// TIA Portal project "FillingLine" (V21)

(* hardware
DEVICE "PLC_Line"  S7-1500 station
   slot 0: "Rail_0"  Rack  6ES7 590-1***0-0AA0
   slot 1: "PLC_Line"  CPU 1516-3 PN/DP  6ES7 516-3AN02-0AB0  V2.9
      slot 3: "CPU display_1"  6ES7591-1BA00-0AA0
      slot 32768: "PROFINET interface_1"  X1
         slot 32769: "Port_1"  X1 P1
         slot 32770: "Port_2"  X1 P2
      slot 33024: "PROFINET interface_2"  X2
         slot 33025: "Port_1"  X2 P1
      slot 33280: "DP interface_1"  X3
      slot 34817: "Virtual CP interface port_1"  Virtual CP interface port  Virtual CP interface port
*)

// ===== PLC "PLC_Line"  CPU 1516-3 PN/DP =====

VAR_GLOBAL   // PLC tag table "Inputs"
   "Button_Start" AT %I0.0 : Bool;   // Start the line
   "Button_Stop" AT %I0.1 : Bool;   // Stop the line, normally closed
   "Button_Reset" AT %I0.2 : Bool;   // Acknowledge faults
   "Infeed_BottleAtFiller" AT %I1.0 : Bool;   // Photo eye: a bottle stands under the filler
   "Infeed_MotorFeedback" AT %I1.1 : Bool;   // Infeed contactor is closed
   "Outfeed_BottleAtEnd" AT %I1.2 : Bool;   // Photo eye at the end of the outfeed
   "Outfeed_MotorFeedback" AT %I1.3 : Bool;   // Outfeed contactor is closed
   "Filler_ValveOpened" AT %I1.4 : Bool;   // Fill valve is open
   "Filler_ValveClosed" AT %I1.5 : Bool;   // Fill valve is closed
   "Packer_Ready" AT %I1.6 : Bool;   // The packer can take a bottle
   "Filler_Level" AT %IW64 : Int;   // Level in the bottle, raw 0 to 27648
END_VAR

VAR_GLOBAL   // PLC tag table "Operator"
   "Recipe_Selected" AT %MW10 : Int;   // Recipe chosen on the panel, 1 to 3
   "Bottles_Filled" AT %MD12 : DInt;   // Bottles filled since the last start
END_VAR

VAR_GLOBAL   // PLC tag table "Outputs"
   "Infeed_Motor" AT %Q0.0 : Bool;   // Infeed conveyor motor
   "Outfeed_Motor" AT %Q0.1 : Bool;   // Outfeed conveyor motor
   "Filler_Valve" AT %Q0.2 : Bool;   // Opens the fill valve
   "Lamp_Running" AT %Q0.3 : Bool;   // The line runs
   "Lamp_Fault" AT %Q0.4 : Bool;   // A fault waits to be acknowledged
END_VAR

// folder: Line

TYPE "typeRecipe"
   STRUCT
      label : String[20];   // Shown on the panel
      volume : Real;   // Fill volume in ml
      settleTime : Time;   // Foam settles before the bottle moves on
   END_STRUCT;
END_TYPE

// folder: Data

DATA_BLOCK "Recipes"   // DB1
{ S7_Optimized_Access := 'TRUE' }
VERSION : 0.1
   VAR
      active : "typeRecipe";   // The recipe in use
      list : Array[1..3] of "typeRecipe";   // Recipes to choose from
   END_VAR
BEGIN
   list[1].label := 'Water 0.5 l';
   list[1].volume := 500.0;
   list[1].settleTime := T#500MS;
   list[2].label := 'Water 1 l';
   list[2].volume := 1000.0;
   list[2].settleTime := T#800MS;
   list[3].label := 'Soda 0.5 l';
   list[3].volume := 480.0;
   list[3].settleTime := T#3S;
END_DATA_BLOCK

DATA_BLOCK "LineData"   // DB2
{ S7_Optimized_Access := 'TRUE' }
VERSION : 0.1
// stored: InstanceOfName FillingLine
"FillingLine"
BEGIN
END_DATA_BLOCK

// folder: (top level)

ORGANIZATION_BLOCK "Main"   // OB1, SCL, ProgramCycle
TITLE = "Main Program Sweep (Cycle)"
{ S7_Optimized_Access := 'TRUE' }
VERSION : 0.1
   VAR_INPUT
      Initial_Call : Bool;   // Initial call of this OB
      Remanence : Bool;   // =True, if remanent data are available
   END_VAR
BEGIN

    // Take the recipe the operator chose, then run the line.
    "Recipes".active := "Recipes".list[LIMIT(MN := 1, IN := "Recipe_Selected", MX := 3)];

    "LineData"(start := "Button_Start",
               stop := NOT "Button_Stop",
               reset := "Button_Reset");

    "Lamp_Running" := "LineData".running;
    "Lamp_Fault" := "LineData".fault;
END_ORGANIZATION_BLOCK

// folder: Common

FUNCTION_BLOCK "Motor"   // FB1, SCL
TITLE = Motor with feedback
{ S7_Optimized_Access := 'TRUE' }
VERSION : 0.1
// Starts and stops a motor and watches its contactor's feedback.
   VAR_INPUT
      start : Bool;   // Start command
      stop : Bool;   // Stop command, wins over start
      feedback : Bool;   // Contactor is closed
      reset : Bool;   // Acknowledge a fault
   END_VAR
   VAR_OUTPUT
      run : Bool;   // Drives the contactor
      fault : Bool;   // The feedback did not come in time
   END_VAR
   VAR
      feedbackTimer : TON_TIME;
      enabled : Bool;   // Started and not stopped since
   END_VAR
   VAR CONSTANT
      FEEDBACK_TIME : Time := T#2S;   // How long the contactor may take
   END_VAR
BEGIN

    // Stop wins over start, and a fault keeps the motor off until it is reset.
    IF #stop OR #fault THEN
        #enabled := FALSE;
    ELSIF #start THEN
        #enabled := TRUE;
    END_IF;

    #feedbackTimer(IN := #enabled AND NOT #feedback,
                   PT := #FEEDBACK_TIME);
    IF #feedbackTimer.Q THEN
        #fault := TRUE;
    ELSIF #reset THEN
        #fault := FALSE;
    END_IF;

    #run := #enabled AND NOT #fault;
END_FUNCTION_BLOCK

FUNCTION_BLOCK "Valve"   // FB2, SCL
TITLE = Valve with end switches
{ S7_Optimized_Access := 'TRUE' }
VERSION : 0.1
// Opens and closes a valve and checks that it reaches its end position in time.
   VAR_INPUT
      open : Bool;   // Open the valve
      opened : Bool;   // End switch: open
      closed : Bool;   // End switch: closed
      reset : Bool;   // Acknowledge a fault
   END_VAR
   VAR_OUTPUT
      output : Bool;   // Drives the valve
      fault : Bool;   // An end position was not reached in time
   END_VAR
   VAR
      moveTimer : TON_TIME;
   END_VAR
   VAR CONSTANT
      MOVE_TIME : Time := T#1S;   // How long the valve may take to move
   END_VAR
BEGIN

    #output := #open AND NOT #fault;

    // The valve is moving while it is not where it was told to go.
    #moveTimer(IN := (#output AND NOT #opened) OR (NOT #output AND NOT #closed),
               PT := #MOVE_TIME);
    IF #moveTimer.Q THEN
        #fault := TRUE;
    ELSIF #reset THEN
        #fault := FALSE;
    END_IF;
END_FUNCTION_BLOCK

FUNCTION "Scale" : Real   // FC1, SCL
TITLE = Scale an analog value
{ S7_Optimized_Access := 'TRUE' }
VERSION : 0.1
// Scales the raw value of an analog input, 0 to 27648, to a range in engineering units.
   VAR_INPUT
      raw : Int;   // Raw value of the analog input
      low : Real;   // Value at 0
      high : Real;   // Value at 27648
   END_VAR
BEGIN

    #Scale := #low + INT_TO_REAL(#raw) / 27648.0 * (#high - #low);
END_FUNCTION

// folder: Line

FUNCTION_BLOCK "Conveyor"   // FB3, SCL
TITLE = Conveyor that holds a bottle at its end
{ S7_Optimized_Access := 'TRUE' }
VERSION : 0.1
// Runs a belt, and stops it while a bottle waits at the end for the next station.
   VAR_INPUT
      enable : Bool;   // The line runs
      bottleAtEnd : Bool;   // Photo eye at the end of the belt
      nextReady : Bool;   // The next station can take the bottle
      motorFeedback : Bool;   // Contactor is closed
      reset : Bool;   // Acknowledge a fault
   END_VAR
   VAR_OUTPUT
      motorOn : Bool;   // Drives the motor
      fault : Bool;   // The motor has a fault
   END_VAR
   VAR
      drive : "Motor";   // The belt's motor
   END_VAR
BEGIN

    // A bottle at the end waits until the next station is ready for it.
    #drive(start := #enable AND (NOT #bottleAtEnd OR #nextReady),
           stop := NOT #enable OR (#bottleAtEnd AND NOT #nextReady),
           feedback := #motorFeedback,
           reset := #reset);

    #motorOn := #drive.run;
    #fault := #drive.fault;
END_FUNCTION_BLOCK

FUNCTION_BLOCK "Filler"   // FB4, SCL
TITLE = Fills one bottle
{ S7_Optimized_Access := 'TRUE' }
VERSION : 0.1
// Fills the bottle under the valve to the recipe's volume, then lets the foam settle.
   VAR_INPUT
      start : Bool;   // A bottle stands under the filler
      levelRaw : Int;   // Level sensor, raw
      valveOpened : Bool;   // End switch: open
      valveClosed : Bool;   // End switch: closed
      recipe : "typeRecipe";   // What to fill
      reset : Bool;   // Acknowledge a fault
   END_VAR
   VAR_OUTPUT
      openValve : Bool;   // Drives the fill valve
      done : Bool;   // The bottle is full and may move on
      fault : Bool;   // The valve has a fault
   END_VAR
   VAR
      "step" : Int;   // 0 idle, 10 filling, 20 settling, 30 done
      level : Real;   // Level in ml
      valve : "Valve";   // The fill valve
      settleTimer : TON_TIME;
   END_VAR
BEGIN

    #level := "Scale"(raw := #levelRaw, low := 0.0, high := 1000.0);

    CASE #step OF
        0:  // Idle: wait for a bottle
            IF #start AND NOT #fault THEN
                #step := 10;
            END_IF;
        10: // Filling: until the recipe's volume is reached
            IF #level >= #recipe.volume THEN
                #step := 20;
            END_IF;
        20: // Settling: the foam goes down
            IF #settleTimer.Q THEN
                #step := 30;
            END_IF;
        30: // Done: wait until the bottle has left
            IF NOT #start THEN
                #step := 0;
            END_IF;
    END_CASE;

    #settleTimer(IN := #step = 20,
                 PT := #recipe.settleTime);
    #valve(open := #step = 10,
           opened := #valveOpened,
           closed := #valveClosed,
           reset := #reset);

    #openValve := #valve.output;
    #done := #step = 30;
    #fault := #valve.fault;
END_FUNCTION_BLOCK

FUNCTION_BLOCK "FillingLine"   // FB5, SCL
TITLE = The filling line
{ S7_Optimized_Access := 'TRUE' }
VERSION : 0.1
// Infeed conveyor, filler and outfeed conveyor, started and stopped as one line.
   VAR_INPUT
      start : Bool;   // Start the line
      stop : Bool;   // Stop the line
      reset : Bool;   // Acknowledge faults
   END_VAR
   VAR_OUTPUT
      running : Bool;   // The line runs
      fault : Bool;   // A station has a fault
   END_VAR
   VAR
      infeed : "Conveyor";   // Brings bottles to the filler
      filler : "Filler";   // Fills them
      outfeed : "Conveyor";   // Takes them to the packer
      lastDone : Bool;   // The filler was done in the last cycle
   END_VAR
BEGIN

    // A fault stops the whole line.
    IF #stop OR #fault THEN
        #running := FALSE;
    ELSIF #start THEN
        #running := TRUE;
        "Bottles_Filled" := 0;
    END_IF;

    // The infeed holds each bottle under the filler until it is full.
    #infeed(enable := #running,
            bottleAtEnd := "Infeed_BottleAtFiller",
            nextReady := #filler.done,
            motorFeedback := "Infeed_MotorFeedback",
            reset := #reset);

    #filler(start := "Infeed_BottleAtFiller" AND #running,
            levelRaw := "Filler_Level",
            valveOpened := "Filler_ValveOpened",
            valveClosed := "Filler_ValveClosed",
            recipe := "Recipes".active,
            reset := #reset);

    #outfeed(enable := #running,
             bottleAtEnd := "Outfeed_BottleAtEnd",
             nextReady := "Packer_Ready",
             motorFeedback := "Outfeed_MotorFeedback",
             reset := #reset);

    // Count each bottle once, when it is done.
    IF #filler.done AND NOT #lastDone THEN
        "Bottles_Filled" := "Bottles_Filled" + 1;
    END_IF;
    #lastDone := #filler.done;

    "Infeed_Motor" := #infeed.motorOn;
    "Outfeed_Motor" := #outfeed.motorOn;
    "Filler_Valve" := #filler.openValve;
    #fault := #infeed.fault OR #filler.fault OR #outfeed.fault;
END_FUNCTION_BLOCK